// TIA Portal V21 export
// export: Created 2026-10-14T03:09:03.7982512Z, ExportSetting WithDefaults, DisplayName Totally Integrated Automation Portal, DisplayVersion V21, DisplayName STEP 7 Professional, DisplayVersion V21, DisplayName STEP 7 Safety, DisplayVersion V21, DisplayName Tech WebApplication, DisplayVersion V21, DisplayName WinCC Basic/Comfort/Advanced, DisplayVersion V21, DisplayName WinCC Unified, DisplayVersion V21
Screen "30_Diagnostics"  800x480, Number=1, Template=01_One_Nav_Level
  on GenerateScreen: SetTag(Tag := MainNavigationState, Value := 3)
  ScreenLayer 
  ScreenLayer 
    GraphicView "Graphic view_2" at 0,0 size 800x480  Picture=PopUpBackground
      VisibilityAnimation "VisibilityAnimation"  RangeEnd=1, RangeStart=1
        tag PopUpBackground
